FUNCTION_BLOCK FB_PulseInterval
VAR_INPUT
	bOn			:	BOOL	:=	FALSE;
	nInterval	:	UDINT	:=	100;		// (Rising edge ~ Rising edge, [ms]) Must be multiple of 20
END_VAR
VAR_OUTPUT
END_VAR
VAR
	nClk		:	UDINT	:=	0;
END_VAR

IF	bOn	THEN
	IF nClk	= 0	THEN
		ExtPort.EL2124_OUT[0]	:=	NOT ExtPort.EL2124_OUT[0];
	END_IF
	IF nClk < TO_UDINT(nInterval / (2 * 10)) THEN
		nClk	:=	nClk + 1;
	ELSE		
		nClk	:=	0;
	END_IF
ELSE
	nClk	:=	0;
	ExtPort.EL2124_OUT[0]	:=	FALSE;
END_IF

END_FUNCTION_BLOCK

(* stored: Version 1.1.0.1, ProductVersion 3.1.4024.15
   POU FB_PulseInterval: Id {4917a029-025d-49c7-9ed5-6eeef52e908a}, SpecialFunc None *)
